TYPE "ST_SequenceCommandLease"
VERSION : 0.1
   STRUCT
      "OwnerIndex" : DInt;
      "ChainIndex" : DInt;
      "Step" : DInt;
      "Raised" : Bool;
      "AbortIssued" : Bool;
      "ReleasedScan" : UDInt;
   END_STRUCT;
END_TYPE
